{attribute 'qualified_only'}
{attribute 'strict'}
TYPE E_CIP_Client_Command :
(
	eDrain := 0,
	eCIP,
	eClose
);
END_TYPE

(* stored: Version 1.1.0.1, ProductVersion 3.1.4024.15
   DUT E_CIP_Client_Command: Id {b3fc0f8e-675a-4a0d-aefe-ed6d65503d84} *)
